TYPE E_MqttLifecyclePhase :
(
    Disconnected,
    OfflineFence,
    Discovery,
    StateSnapshot,
    OnlineAnnouncement,
    Ready
);
END_TYPE

(* stored: Version 1.1.0.1
   DUT E_MqttLifecyclePhase: Id {75c6111c-20ce-4ed4-b451-1f722f4d1409} *)
